FUNCTION F_NumericObjectPool_S_TO_OBJID (* Extract the ISOBUS Object ID (u16ObjId) out of a NumericObjectPool_S struct. *)
  (* Standard: 61499-2; Description: Copyright (c) 2026 Meisterschulen am Ostbahnhof This program and the accompanying materials are made available under the terms of the Eclipse Public License 2.0 which is available at https://www.eclipse.org/legal/epl-2.0/ SPDX-License-Identifier: EPL-2.0 *)
  (* Version 1.0, 2026-10-11, Franz Höpfinger, Meisterschulen am Ostbahnhof *)
  PACKAGE logiBUS::utils::conversion::phys;
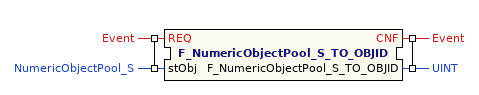
  EVENT_INPUT
    REQ WITH stObj;
  END_EVENT
  EVENT_OUTPUT
    CNF WITH F_NumericObjectPool_S_TO_OBJID;
  END_EVENT
  VAR_INPUT
    stObj : logiBUS::utils::conversion::phys::NumericObjectPool_S;
  END_VAR
  VAR_OUTPUT
    F_NumericObjectPool_S_TO_OBJID : UINT;
  END_VAR
  BODY IN ST:
PACKAGE logiBUS::utils::conversion::phys;

(* Extract the ISOBUS Object ID (u16ObjId) out of a NumericObjectPool_S struct. *)
FUNCTION F_NumericObjectPool_S_TO_OBJID : UINT

VAR_INPUT
	stObj : NumericObjectPool_S;
END_VAR

F_NumericObjectPool_S_TO_OBJID := stObj.u16ObjId;

END_FUNCTION
  END_BODY
END_FUNCTION
